Staubli VAL3: safeLogic.pjx

--- safeLogic.pjx ---
Parameters version=s8.12.1Cs9_BS2449 stackSize=5000 millimeterUnit=true
Program file=areaCheck.pgx
Program file=checkPoint.pgx
Program file=computeArea.pgx
Program file=loadLib.pgx
Program file=main.pgx
Program file=start.pgx
Program file=stop.pgx
Data file=safeLogic.dtx
Library alias=safeData path=Disk://data/CustomerLib/default/safeData/safeData.pjx
Library alias=rs path=Disk://source/projectSource/robotStatus/robotStatus.pjx
Library alias=saveData path=Disk://source/saveData/saveData.pjx
Library alias=io path=Disk://source/projectSource/io/io.pjx

--- safeLogic.dtx ---
mdesc mNomSpeed
num nLastLib

--- main.pgx ---
public program main()
  local pointRx l_pPoint
  local num l_nResult
  local tool l_tTool
begin
  //  nLastLib=-1
  do
//    call saveData:getTool(saveData:nJogTool,l_tTool)
//    l_pPoint=here(l_tTool,world)

    call areaCheck()
    call checkPoint()


    delay(0)
  until false

end

--- start.pgx ---
program start()
begin
end

--- areaCheck.pgx ---
public program areaCheck()
  local num l_i
begin
  for l_i = 0 to size(safeData:zZoneItem)-1
    if safeData:zZoneItem[l_i].bActive
      call computeArea(l_i)
    endIf
  endFor

end

--- checkPoint.pgx ---
public program checkPoint()
  local num l_nSize
  local num l_i
  local pointRx l_pPoint
  local bool l_bErr
begin
  l_pPoint=here(flange,world)
  l_nSize=size(safeData:sSPoint)
  for l_i = 0 to l_nSize-1
    if safeData:sSPoint[l_i].bActive
      if distance(safeData:sSPoint[l_i].pPointRx.trsf,l_pPoint.trsf)<5
        call io:setDigOutput(io:dOutput[l_i+96],true,l_bErr)
      else
        call io:setDigOutput(io:dOutput[l_i+96],false,l_bErr)
      endIf
    endIf
  endFor
end

--- computeArea.pgx ---
public program computeArea(num x_nIndex)
  local trsf l_trsf1
  local trsf l_trsf2
  local num l_nMinX
  local num l_nMinY
  local num l_nMinZ
  local num l_nMaxX
  local num l_nMaxY
  local num l_nMaxZ
  local bool l_bResult
  local bool l_bResult1
  local bool l_bResult2
  local bool l_bErr
  local frame l_fFrame
  local pointRx l_pPoint
  local tool l_tTool
begin

  link(l_pPoint,l_fFrame)
  link(l_fFrame,world)
  l_fFrame.trsf=safeData:zZoneItem[x_nIndex].fBase.trsf


  call saveData:getTool(saveData:nJogTool,l_tTool)
  l_pPoint=here(l_tTool,l_fFrame)


  l_trsf1.x=safeData:zZoneItem[x_nIndex].pFirst.trsf.x
  l_trsf1.y=safeData:zZoneItem[x_nIndex].pFirst.trsf.y
  l_trsf1.z=safeData:zZoneItem[x_nIndex].pFirst.trsf.z

  l_trsf2.x=l_trsf1.x+safeData:zZoneItem[x_nIndex].pSecond.trsf.x
  l_trsf2.y=l_trsf1.y+safeData:zZoneItem[x_nIndex].pSecond.trsf.y
  l_trsf2.z=l_trsf1.z+safeData:zZoneItem[x_nIndex].pSecond.trsf.z

  l_nMinX=min(l_trsf1.x,l_trsf2.x)
  l_nMinY=min(l_trsf1.y,l_trsf2.y)
  l_nMinZ=min(l_trsf1.z,l_trsf2.z)
  l_nMaxX=max(l_trsf1.x,l_trsf2.x)
  l_nMaxY=max(l_trsf1.y,l_trsf2.y)
  l_nMaxZ=max(l_trsf1.z,l_trsf2.z)

  if l_nMinX<=l_pPoint.trsf.x and l_pPoint.trsf.x<=l_nMaxX
    l_bResult=true
  else
    l_bResult=false
  endIf
  if l_nMinY<=l_pPoint.trsf.y and l_pPoint.trsf.y<=l_nMaxY
    l_bResult1=true
  else
    l_bResult1=false
  endIf
  if l_nMinZ<=l_pPoint.trsf.z and l_pPoint.trsf.z<=l_nMaxZ
    l_bResult2=true
  else
    l_bResult2=false
  endIf
  //如果是=0，不发送信号（0不起作用）
  if l_bResult and l_bResult1 and l_bResult2
    call io:setDigOutput(io:dOutput[x_nIndex+112],true,l_bErr)
  else
    call io:setDigOutput(io:dOutput[x_nIndex+112],false,l_bErr)
  endIf
end

--- loadLib.pgx ---
public program loadLib(num x_nLib, num& x_nResult)
  local string l_sPath
begin
  if x_nLib>=0
    l_sPath="Disk://data/CustomerLib/lib"+toString("",x_nLib)+"/safeData"
    x_nResult=safeData:libLoad(l_sPath)
    wait(x_nResult==0)
  else
    call rs:setAlarm(302,0)
  endIf
end

--- stop.pgx ---
program stop()
begin
end
